// TIA Portal V21 export
TagTable "T_V8"
  Y_V8 : USInt  (PLC tag HMI_IF.State, HMI_Connection_1, 1 s)
